Fanuc KAREL source: KT00539.KL

PROGRAM KT00539
%NOLOCKGROUP
VAR
  P1: JOINTPOS
  P2: XYZWPR
  OUT: POSITION
BEGIN
    P2.Y = 2.0
  OUT = P1 : P2
END KT00539
